// TIA Portal V21 export
FUNCTION "F_FC_Logic" : Void   // FC9, F_FBD
{ S7_Optimized_Access := 'TRUE' }
   VAR_INPUT
      GuardClosed : Bool;   // Schutztür geschlossen / Guard door closed
      SetupMode : Bool;   // Einrichtbetrieb angewählt / Setup mode selected
      EmergencyStopOk : Bool;   // Not-Halt nicht betätigt / Emergency stop not pressed
   END_VAR
   VAR_OUTPUT
      Release : Bool;   // Freigabe der Maschine / Release of the machine
   END_VAR
BEGIN

REGION Network 1: Schutztür oder Einrichtbetrieb, und Not-Halt in Ordnung / Guard or setup mode, and emergency stop ok
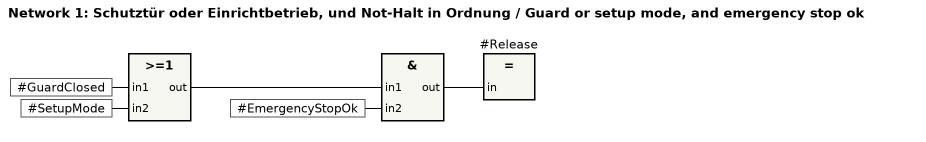
   #Release := (#GuardClosed OR #SetupMode) AND #EmergencyStopOk;
END_REGION
END_FUNCTION
